(* Logix 5000 project; controller DSFW_Budzar vendor 1 type 14 code 154 rev 32.13; software revision 32.03; part 5 of 5 *)
(* tags used below, declared in another part *)
   Active_Setpoint : REAL;
   Batch_Mode_Enable : BOOL;
   FCV_101 : ALIAS FOR Local:8:O.Ch2Data;   // Process Bypass Flow Control Valve
   FIC_101_Manual_Percent : REAL;
   FIC_101_Run_PID : BOOL;
   FIC_101_Setpoint : REAL;
   FIC_101_Stop_PID : BOOL;
   FIT_101 : BL_Analog_Input;   // Flow Indicating Transmitter
   FIT_101_PID_Scale_Max : REAL;
   FIT_101_PID_Scale_Min : REAL;
   HMI_FCV_101_CV : REAL;
   HMI_FCV_101_Lamp : BOOL;
   HMI_PCV_101_Lamp : BOOL;
   HMI_PCV_101_Output : REAL;
   PCV_101_Auto_Manual : BOOL;
   PCV_101_Flush_Position : REAL;   // PCV-101 Desired Flush Position (4000-20000 counts)
   PCV_101_Manual_Output : REAL;
   PCV_101_Multiplexer : DINT;   // Selects controlling input to multiplxer
   PCV_101_Pressure_SP : REAL;
   PCV_101_Run_PIDE : BOOL;
   PCV_101_Start_Position : REAL;   // PCV-101 Desired Start Position (4000-20000 counts)
   PCV_101_Stop_PIDE : BOOL;
   PT_103 : BL_Analog_Input;   // R404A Compressor Discharge Pressure
   PT_103_PID_Scale_Max : REAL;
   PT_103_PID_Scale_Min : REAL;
   PT_104 : BL_Analog_Input;   // R404A Evaporator Suction Pressure
   Ramp_Soak_Segments_HMI_Set : REAL;
   REACTOR_BATCH_PID_START : BOOL;
   REACTOR_BATCH_PID_STOP : BOOL;
   REACTOR_BATCH_PIDE_CV_AS_SP : REAL;
   REACTOR_BATCH_PV : REAL;
   REACTOR_HEAT_RUN_PIDE : BOOL;
   REACTOR_HEAT_STOP_PIDE : BOOL;
   RX_RMPS_Output : REAL;
   RX_RMPS_Ramp_Value : REAL[11];
   RX_RMPS_Soak_Time : REAL[11];
   RX_RMPS_Soak_Value : REAL[11];
   RX_RMPS_SP_Out : REAL;
   RX_Run_Temp_Profile : BOOL;
   RX_Start_Temperature_Profile : BOOL;
   RX_Stop_Temp_Profile : BOOL;
   SCR_101_Auto_Manual : BOOL;
   SCR_101_Manual_Output : REAL;
   SCR_PID_Request : REAL;
   TCV_101_Auto_Manual : BOOL;
   TCV_101_Manual_Output : REAL;
   TCV_101_Pressure_Setpoint : REAL;   // TCV-101 Hot Gas Pressure PID loop Setpoint
   TCV_101_Run_PIDE : BOOL;
   TCV_101_Stop_PIDE : BOOL;
   TCV_CV : REAL;   // TCV Loop Output Scaled (0-100%)
   TCV_Multiplexer : DINT;
   TE_101 : BL_Analog_Input;   // Process Supply Temperature
   Temperature_Setpoint : REAL;
   VESSEL_TEMPERATURE : BL_Analog_Input;   // End User Reactor Temperature
(* EEV_PID, continued *)

ROUTINE Routine_Schedule   (* ladder *)
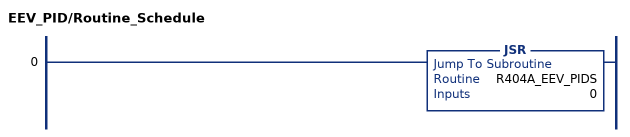
   0: JSR(R404A_EEV_PIDS,0);
END_ROUTINE
END_PROGRAM

PROGRAM Main   (* main routine Routine_Schedule *)
VAR
   ADD_01 : FBD_MATH := (SourceA := 5.0, SourceB := 1.0, Dest := 6.0);
   BOR_01 : FBD_BOOLEAN_OR;
   BOR_02 : FBD_BOOLEAN_OR;
   ESEL_03 : SELECT_ENHANCED := (In1 := 4000.0, In2 := 4000.0, InsUsed := 2, SelectorMode := 1, OperSelector := 1, ProgProgReq := 1, Out := 4000.0, SelectedIn := 1, ProgOper := 1);
   GEQ_02 : FBD_COMPARE := (SourceB := 0.5);
   MUX_01 : MULTIPLEXER := (In1 := 4000.0, In2 := 4000.0, In3 := 8800.0, Selector := 1, Out := 4000.0);
   PIDE_01 : PID_ENHANCED := (PVEUMax := 140.0, SPProg := 20.0, SPHLimit := 125.0, RatioProg := 1.0, RatioOper := 1.0, RatioHLimit := 1.0, RatioLLimit := 1.0, CVEUMax := 100.0, CVHLimit := 100.0, ControlAction := 1, PGain := 2.0, IGain := 1.0, PVEDerivative := 1, DSmoothing := 1, PVTracking := 1, ProgOverrideReq := 1, RTSTime := 1, InitPrimary := 1, Ratio := 1.0, Override := 1, DeltaT := 0.1);
   SCL_05 : SCALE := (In := 4000.0, InRawMax := 20000.0, InRawMin := 4000.0, InEUMax := 100.0);
   SEL_01 : SELECT := (In1 := 6590.2725, In2 := 12000.0, Out := 6590.2725);
   SEL_02 : SELECT;
   SEL_03 : SELECT := (In1 := 23.3, In2 := 20.0, Out := 23.3);
   SEL_04 : SELECT := (In1 := 20.0, In2 := 20.0, Out := 20.0);
   SEL_09 : SELECT := (In1 := 4000.0, In2 := 4000.0, Out := 4000.0);
END_VAR

ROUTINE Process_PIDS   (* function block diagram *)
   SHEET 1
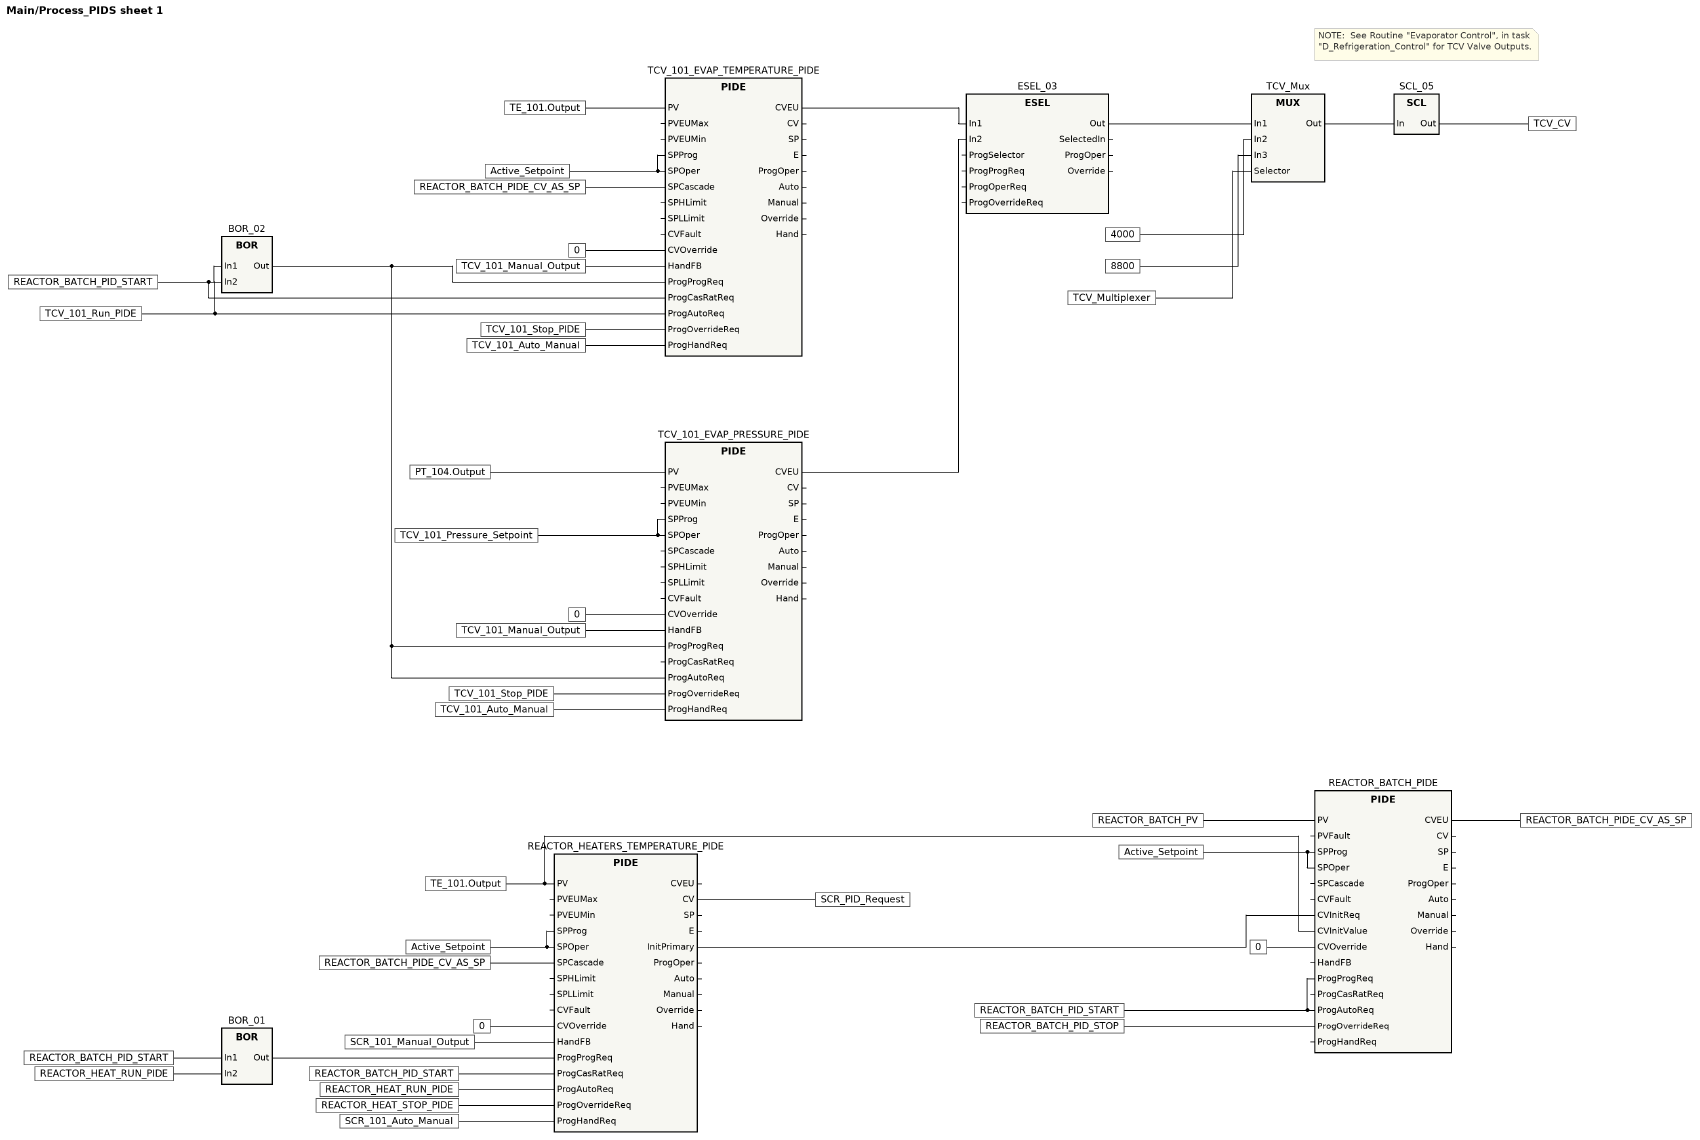
   // NOTE:  See Routine "Evaporator Control", in task "D_Refrigeration_Control" for TCV Valve Outputs.
   BOR_02 : BOR(In1 := REACTOR_BATCH_PID_START, In2 := TCV_101_Run_PIDE);
   BOR_01 : BOR(In1 := REACTOR_BATCH_PID_START, In2 := REACTOR_HEAT_RUN_PIDE);
   REACTOR_HEATERS_TEMPERATURE_PIDE : PIDE(PV := TE_101.Output, SPProg := Active_Setpoint, SPOper := Active_Setpoint, SPCascade := REACTOR_BATCH_PIDE_CV_AS_SP, CVOverride := 0, HandFB := SCR_101_Manual_Output, ProgProgReq := BOR_01.Out, ProgCasRatReq := REACTOR_BATCH_PID_START, ProgAutoReq := REACTOR_HEAT_RUN_PIDE, ProgOverrideReq := REACTOR_HEAT_STOP_PIDE, ProgHandReq := SCR_101_Auto_Manual);   // unwired pins: PVEUMax PVEUMin SPHLimit SPLLimit CVFault CVEU SP E ProgOper Auto Manual Override Hand
   TCV_101_EVAP_TEMPERATURE_PIDE : PIDE(PV := TE_101.Output, SPProg := Active_Setpoint, SPOper := Active_Setpoint, SPCascade := REACTOR_BATCH_PIDE_CV_AS_SP, CVOverride := 0, HandFB := TCV_101_Manual_Output, ProgProgReq := BOR_02.Out, ProgCasRatReq := REACTOR_BATCH_PID_START, ProgAutoReq := TCV_101_Run_PIDE, ProgOverrideReq := TCV_101_Stop_PIDE, ProgHandReq := TCV_101_Auto_Manual);   // unwired pins: PVEUMax PVEUMin SPHLimit SPLLimit CVFault CV SP E ProgOper Auto Manual Override Hand
   TCV_101_EVAP_PRESSURE_PIDE : PIDE(PV := PT_104.Output, SPProg := TCV_101_Pressure_Setpoint, SPOper := TCV_101_Pressure_Setpoint, CVOverride := 0, HandFB := TCV_101_Manual_Output, ProgProgReq := BOR_02.Out, ProgAutoReq := BOR_02.Out, ProgOverrideReq := TCV_101_Stop_PIDE, ProgHandReq := TCV_101_Auto_Manual);   // unwired pins: PVEUMax PVEUMin SPCascade SPHLimit SPLLimit CVFault ProgCasRatReq CV SP E ProgOper Auto Manual Override Hand
   SCR_PID_Request := REACTOR_HEATERS_TEMPERATURE_PIDE.CV;
   ESEL_03 : ESEL(In1 := TCV_101_EVAP_TEMPERATURE_PIDE.CVEU, In2 := TCV_101_EVAP_PRESSURE_PIDE.CVEU);   // unwired pins: ProgSelector ProgProgReq ProgOperReq ProgOverrideReq SelectedIn ProgOper Override
   TCV_Mux : MUX(In1 := ESEL_03.Out, In2 := 4000, In3 := 8800, Selector := TCV_Multiplexer);
   REACTOR_BATCH_PIDE : PIDE(PV := REACTOR_BATCH_PV, SPProg := Active_Setpoint, SPOper := Active_Setpoint, CVInitReq := REACTOR_HEATERS_TEMPERATURE_PIDE.InitPrimary, CVInitValue := TE_101.Output, CVOverride := 0, ProgProgReq := REACTOR_BATCH_PID_START, ProgAutoReq := REACTOR_BATCH_PID_START, ProgOverrideReq := REACTOR_BATCH_PID_STOP);   // unwired pins: PVFault SPCascade CVFault HandFB ProgCasRatReq ProgHandReq CV SP E ProgOper Auto Manual Override Hand
   SCL_05 : SCL(In := TCV_Mux.Out);
   REACTOR_BATCH_PIDE_CV_AS_SP := REACTOR_BATCH_PIDE.CVEU;
   TCV_CV := SCL_05.Out;
END_ROUTINE

ROUTINE RMPS   (* function block diagram *)
   SHEET 1
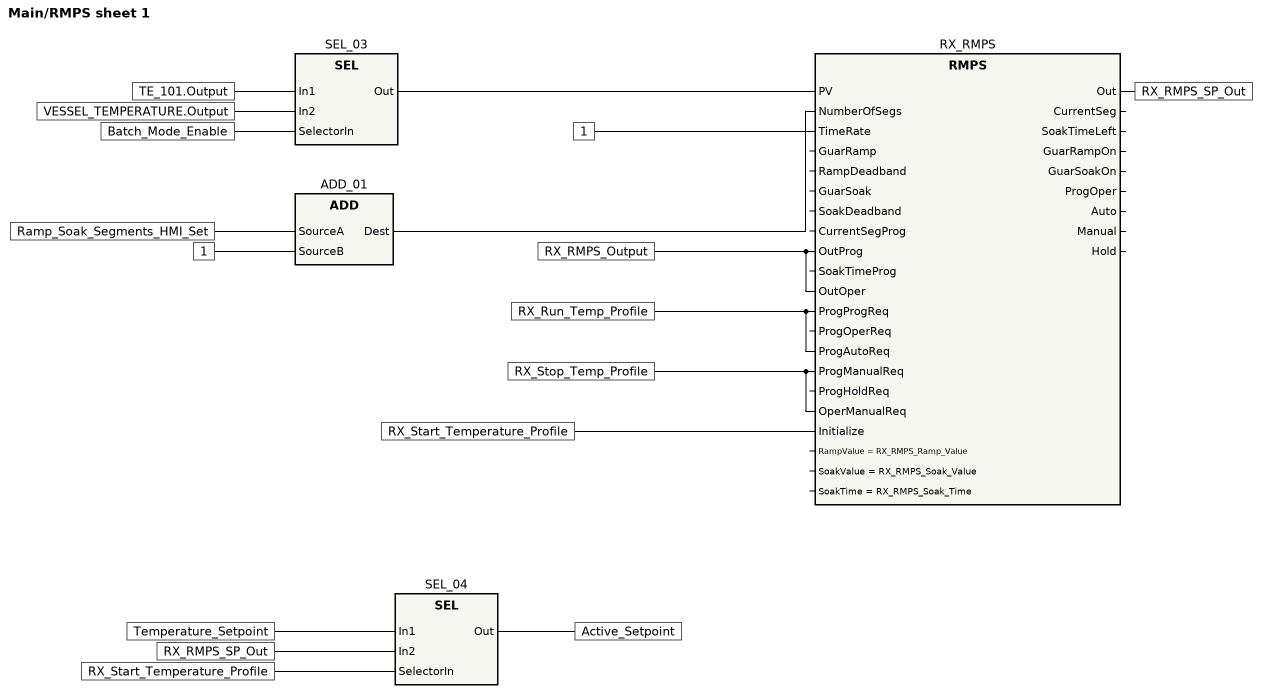
   SEL_03 : SEL(In1 := TE_101.Output, In2 := VESSEL_TEMPERATURE.Output, SelectorIn := Batch_Mode_Enable);
   ADD_01 : ADD(SourceA := Ramp_Soak_Segments_HMI_Set, SourceB := 1);
   SEL_04 : SEL(In1 := Temperature_Setpoint, In2 := RX_RMPS_SP_Out, SelectorIn := RX_Start_Temperature_Profile);
   Active_Setpoint := SEL_04.Out;
   RX_RMPS : RMPS(PV := SEL_03.Out, NumberOfSegs := ADD_01.Dest, TimeRate := 1, OutProg := RX_RMPS_Output, OutOper := RX_RMPS_Output, ProgProgReq := RX_Run_Temp_Profile, ProgAutoReq := RX_Run_Temp_Profile, ProgManualReq := RX_Stop_Temp_Profile, OperManualReq := RX_Stop_Temp_Profile, Initialize := RX_Start_Temperature_Profile, RampValue := RX_RMPS_Ramp_Value, SoakValue := RX_RMPS_Soak_Value, SoakTime := RX_RMPS_Soak_Time);   // unwired pins: GuarRamp RampDeadband GuarSoak SoakDeadband CurrentSegProg SoakTimeProg ProgOperReq ProgHoldReq CurrentSeg SoakTimeLeft GuarRampOn GuarSoakOn ProgOper Auto Manual Hold
   RX_RMPS_SP_Out := RX_RMPS.Out;
END_ROUTINE

ROUTINE Routine_Schedule   (* ladder *)
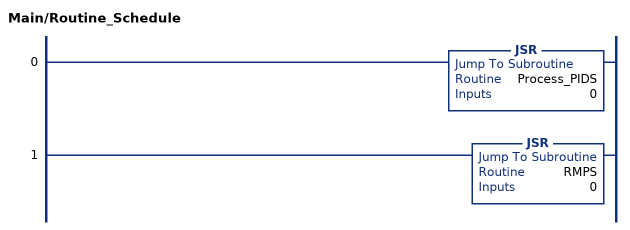
   0: JSR(Process_PIDS,0);
   1: JSR(RMPS,0);
END_ROUTINE
END_PROGRAM

PROGRAM Pressure_PID   (* main routine Routine_Schedule *)
VAR
   GEQ_01 : FBD_COMPARE := (SourceA := 4000.0, SourceB := 0.5, Dest := 1);
   GEQ_02 : FBD_COMPARE := (SourceA := 4000.0, SourceB := 4100.0);
   GEQ_03 : FBD_COMPARE := (SourceB := 4100.0);
   MUX_01 : MULTIPLEXER := (In1 := 4000.0, In2 := 12000.0, In3 := 20000.0, Selector := 1, Out := 4000.0);
   SCL_01 : SCALE := (In := 4000.0, InRawMax := 20000.0, InRawMin := 4000.0, InEUMax := 100.0);
   SCL_02 : SCALE := (In := 4000.0, InRawMax := 20000.0, InRawMin := 4000.0, InEUMax := 100.0);
   SEL_01 : SELECT := (In1 := 4000.0, In2 := 12000.0, Out := 4000.0);
END_VAR

ROUTINE FIC_101   (* function block diagram *)
   SHEET 1
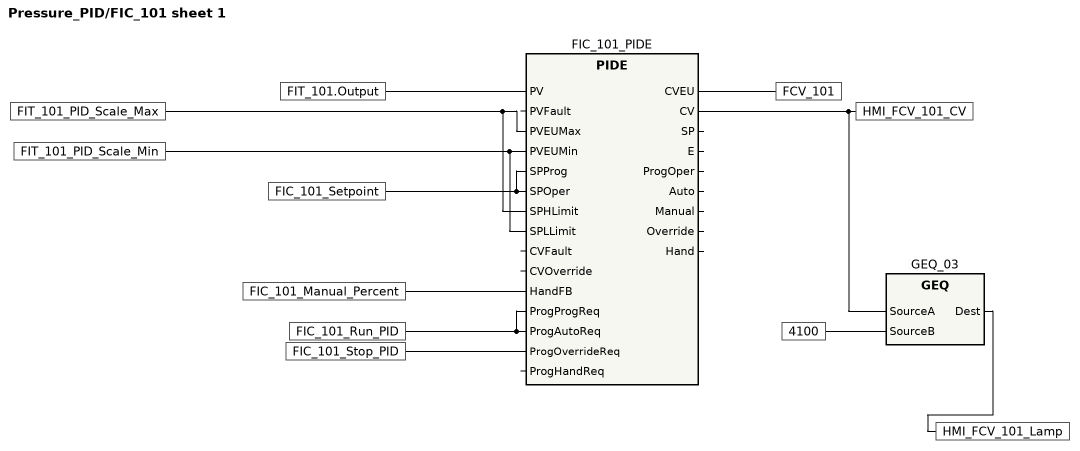
   FIC_101_PIDE : PIDE(PV := FIT_101.Output, PVEUMax := FIT_101_PID_Scale_Max, PVEUMin := FIT_101_PID_Scale_Min, SPProg := FIC_101_Setpoint, SPOper := FIC_101_Setpoint, SPHLimit := FIT_101_PID_Scale_Max, SPLLimit := FIT_101_PID_Scale_Min, HandFB := FIC_101_Manual_Percent, ProgProgReq := FIC_101_Run_PID, ProgAutoReq := FIC_101_Run_PID, ProgOverrideReq := FIC_101_Stop_PID);   // unwired pins: PVFault CVFault CVOverride ProgHandReq SP E ProgOper Auto Manual Override Hand
   FCV_101 := FIC_101_PIDE.CVEU;
   HMI_FCV_101_CV := FIC_101_PIDE.CV;
   GEQ_03 : GEQ(SourceA := FIC_101_PIDE.CV, SourceB := 4100);
   HMI_FCV_101_Lamp := GEQ_03.Dest;
END_ROUTINE

ROUTINE PCV_101   (* function block diagram *)
// Condenser Pressure Control
   SHEET 1
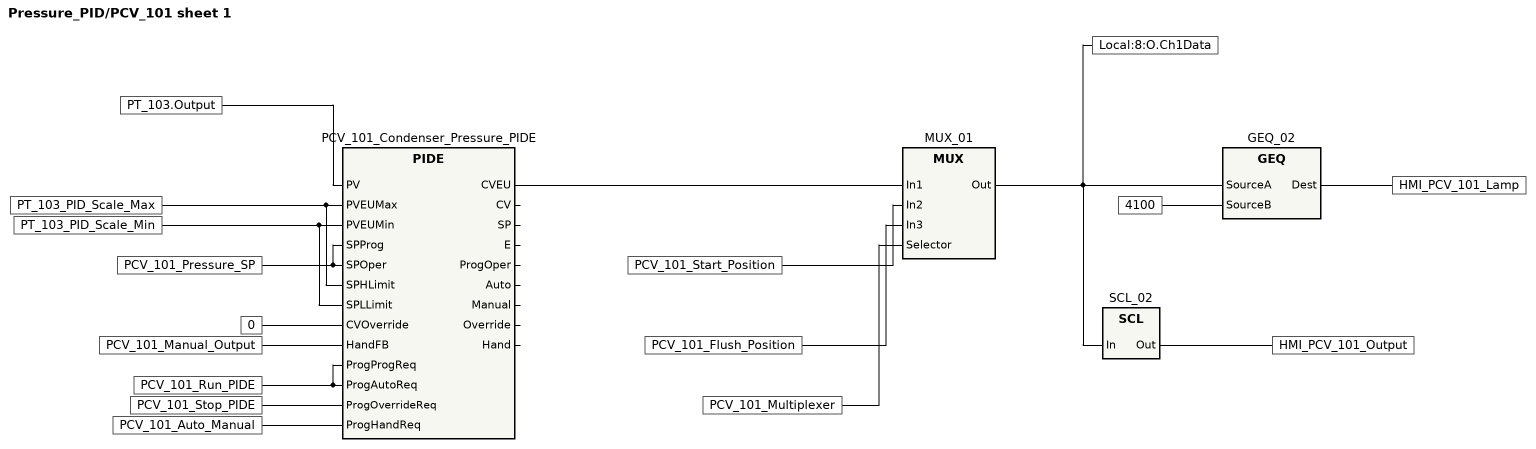
   PCV_101_Condenser_Pressure_PIDE : PIDE(PV := PT_103.Output, PVEUMax := PT_103_PID_Scale_Max, PVEUMin := PT_103_PID_Scale_Min, SPProg := PCV_101_Pressure_SP, SPOper := PCV_101_Pressure_SP, SPHLimit := PT_103_PID_Scale_Max, SPLLimit := PT_103_PID_Scale_Min, CVOverride := 0, HandFB := PCV_101_Manual_Output, ProgProgReq := PCV_101_Run_PIDE, ProgAutoReq := PCV_101_Run_PIDE, ProgOverrideReq := PCV_101_Stop_PIDE, ProgHandReq := PCV_101_Auto_Manual);   // unwired pins: CV SP E ProgOper Auto Manual Override Hand
   MUX_01 : MUX(In1 := PCV_101_Condenser_Pressure_PIDE.CVEU, In2 := PCV_101_Start_Position, In3 := PCV_101_Flush_Position, Selector := PCV_101_Multiplexer);
   Local:8:O.Ch1Data := MUX_01.Out;
   SCL_02 : SCL(In := MUX_01.Out);
   GEQ_02 : GEQ(SourceA := MUX_01.Out, SourceB := 4100);
   HMI_PCV_101_Output := SCL_02.Out;
   HMI_PCV_101_Lamp := GEQ_02.Dest;
END_ROUTINE

ROUTINE Routine_Schedule   (* ladder *)
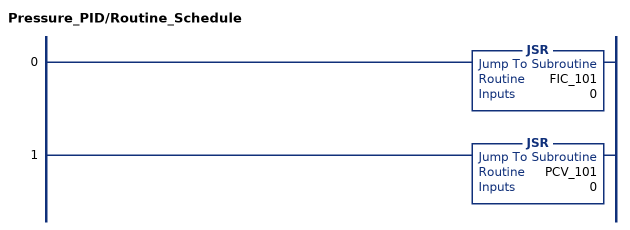
   0: JSR(FIC_101,0);
   1: JSR(PCV_101,0);
END_ROUTINE
END_PROGRAM
